Fanuc KAREL source: KT00881.KL

PROGRAM KT00881
%NOLOCKGROUP
VAR
  I1: INTEGER
  I2: INTEGER
  OUT: REAL
BEGIN
  I1 = 2
  I2 = 3
  I1 = 2
  I2 = 3
  OUT = ATAN2(I1, I1)
END KT00881
